TYPE ET_BECKHOFF_AxisSetLimits :
(
	eWaitExecute := 0,
	eSetReferenceSystem,
	eWfSetReferenceSystem,
	eSetPositionBias,
	eWfSetPositionBias,
	eSetLimitPos,
	eWfSetLimitPos,
	eSetLimitNeg,
	eWfSetLimitNeg,
	eEnableLimitPos,
	eWfEnableLimitPos,
	eEnableLimitNeg,
	eWfEnableLimitNeg,
	eEnablePosLagMonitoring,
	eWfEnablePosLagMonitoring,
	eDone := 197,
	eError := 198,
	eNoExecute := 199
);
END_TYPE

(* stored: Version 1.1.0.1, ProductVersion 3.1.4024.15
   DUT ET_BECKHOFF_AxisSetLimits: Id {f18df66e-840b-4f5a-b718-f8a294d3f82d} *)
